Staubli VAL3: movePoint.pgx

public program movePoint(num x_nIndex)
  local pointRx l_pPoint
  local bool l_bResult
  local tool l_tTool
begin

  l_bResult=userPageConfirm("是否移动到此点位？")

  if l_bResult
    resetMotion()
    link(l_pPoint,fFrame)
    call saveData:getTool(saveData:nJogTool,l_tTool)
    l_pPoint.trsf=safeTemp:zZoneItem[x_nIndex].pFirst.trsf
    l_pPoint.config=safeTemp:zZoneItem[x_nIndex].pFirst.config
    movej(l_pPoint,l_tTool,mNomSpeed)
    delay(0)
  endIf
end
